{region 'Documentation'}
(*!
<summary>Checks whether the USINT value is inside the inclusive range.</summary>
<description>

Minimum &gt; Maximum reports Error during active evaluation; equal bounds are
valid.

</description>
*)
{endregion}
FUNCTION_BLOCK AssertInRange_USInt EXTENDS AssertionBase
VAR_INPUT
    IN : USINT; //! Actual value checked or observed by this Assertion.
    Minimum : USINT; //! Inclusive lower bound of the comparison; for a range, must not exceed Maximum.
    Maximum : USINT; //! Inclusive upper bound of the comparison; for a range, must not be below Minimum.
END_VAR

SUPER^();

{region 'Documentation'}
(*!
<summary>Check whether the USINT value is inside the inclusive range.</summary>
*)
{endregion}
METHOD PROTECTED Assert
VAR
    Message : STRING(GVL_Constants.MessageLength);
    MinimumText : STRING(GVL_Constants.AssertionValueLength);
    MaximumText : STRING(GVL_Constants.AssertionValueLength);
    ActualText : STRING(GVL_Constants.AssertionValueLength);
END_VAR
IF NOT EvaluationActive THEN
    RETURN;
END_IF;

IF Result = E_Result.Error THEN
    RETURN;
END_IF;

IF Minimum > Maximum THEN
    MinimumText := USINT_TO_STRING(Minimum);
    MaximumText := USINT_TO_STRING(Maximum);
    Message := CONCAT('Assertion error: minimum exceeds maximum. Minimum = ',
        MinimumText);
    Message := CONCAT(Message, ', Maximum = ');
    Message := CONCAT(Message, MaximumText);
    Message := CONCAT(Message, '.');
    Error(Message := Message);
    RETURN;
END_IF;

IF Result = E_Result.Failed THEN
    RETURN;
END_IF;

IF (IN < Minimum) OR (IN > Maximum) THEN
    MinimumText := USINT_TO_STRING(Minimum);
    MaximumText := USINT_TO_STRING(Maximum);
    ActualText := USINT_TO_STRING(IN);
    Message := CONCAT('Assertion failed: value is outside allowed range. Minimum = ',
        MinimumText);
    Message := CONCAT(Message, ', Maximum = ');
    Message := CONCAT(Message, MaximumText);
    Message := CONCAT(Message, ', Actual = ');
    Message := CONCAT(Message, ActualText);
    Message := CONCAT(Message, '.');
    Fail(Message := Message);
    RETURN;
END_IF;

Pass();
END_METHOD

END_FUNCTION_BLOCK

(* stored: Version 1.1.0.1
   POU AssertInRange_USInt: Id {109473ef-00d4-4d34-a6d0-0e85c4dd07a7}, SpecialFunc None
   Folder Internal: Id {37c41550-f958-41ee-8485-ee928133fb56}
   Method Assert: Id {15ceaf6b-0212-4032-9e41-417269f15a58} *)
